// TIA Portal V19 export
DATA_BLOCK "iFB_AutoMode"   // DB16
// stored: InstanceOfName FB_AutoMode, InstanceOfType FB
"FB_AutoMode"
   // VAR_INPUT
   //    Enable : Bool;
   //    In_xBatchLoaded : Bool;
   //    In_xPickProductPresent : Bool;
   //    In_ProductConveyor_Pos1 : Bool;
   //    In_ProductConveyor_Pos3 : Bool;
   //    xKillAll : Bool;
   //    In_xPressClosed : Bool;
   //    xProduct_Conv_Exit : Bool;
   //    In_Safety : Bool;
   //    In_ExecuteHomeR1 : Bool;
   //    In_ExecuteHomeR2 : Bool;
   //    In_ExecuteHomeR3 : Bool;
   //    "In_Execute HomeR4" : Bool;
   // END_VAR
   // VAR_IN_OUT
   //    Servo : "ST_Servo";
   //    Robot : Array[1..3] of "ST_ROBOT";
   // END_VAR
   // VAR
   //    "iStage-R1" : Int;
   //    "iStage-R2" : Int;
   //    "iStage-R3" : Int;
   //    "iStage-Press" : Int;
   //    "iStage-Servo" : Int;
   //    xPickR1 : Bool;
   //    xPickR2 : Bool;
   //    xPickR3 : Bool;
   //    xPlaceR1 : Bool;
   //    xPlaceR2 : Bool;
   //    xPlaceR3 : Bool;
   //    xHommingR1 : Bool;
   //    xHommingR2 : Bool;
   //    xHommingR3 : Bool;
   //    xHommingServo : Bool;
   //    xPressEnable : Bool;
   //    xPressCycle : Bool;
   //    Conveyor_Busy : Bool;
   //    Conveyor_Done : Bool;
   //    xProductAtPress : Bool;
   //    xPressProductedReady : Bool;
   //    xServoProductPos1 : Bool;
   //    xServoProductPos2 : Bool;
   //    xServoProductPos3 : Bool;
   //    xServoClearRequest : Bool;
   //    iServoClearStep : Int;
   //    xHomming : Bool;
   // END_VAR
BEGIN
END_DATA_BLOCK
